(* IEC 61131-3 sources: Gen-AI/final/Gen-AI_v1.0_submission/A2_框架源码/agent/logs/full34_fixture/E3_S13_1_42/tools/candidate_1/fixture_compile, 1 file *)

(* ---- source.st ---- *)
FUNCTION_BLOCK FB_S13
VAR_INPUT
    LineRun : BOOL;
    PartAtMerge : BOOL;
    PartOnMain : BOOL;
    JamSensor : BOOL;
    ResetBtn : BOOL;
    ModeAuto : BOOL;
END_VAR
VAR_OUTPUT
    MainMotor : BOOL;
    MergeMotor : BOOL;
    SpeedHigh : BOOL;
    JamAlarm : BOOL;
    Status : WORD;
END_VAR
(* Add a VAR block for internal state/timers before the implementation, if needed. *)
(* SKELETON ONLY: replace this RETURN with scan logic and required initial state. *)
RETURN;
END_FUNCTION_BLOCK

(* FIXTURE_COMPILE_FAIL *)
